Fanuc KAREL source: ko00069.KL

-- PROVISIONAL review KL for V1013-1; original PC SHA256 da2f10e1df383914801fae96bc6c5efdb4d0e3289bffabeefbd34ef2aa823d8f
-- Incomplete behavior may be omitted. Consult companion uncertainty JSON. Do not deploy.
PROGRAM KO00069
%NOLOCKGROUP
BEGIN
  -- UNRESOLVED_PC offsets 5-12; opcodes 9D,23
  -- UNRESOLVED_PC offsets 17-66; opcodes 27,22,1C,27,49,7E,AD,22,31,7E,4A
  -- UNRESOLVED_PC offsets 71-75; opcodes 7F
END KO00069
